Fanuc KAREL source: KB00038.KL

PROGRAM KB00038
%NOLOCKGROUP
VAR
  P1: REAL
  P2: JOINTPOS
  P3: INTEGER
BEGIN
  P1 = 1.0
  P3 = 1
  CNV_REL_JPOS(P1, P2, P3)
END KB00038
